Fanuc KAREL source: KT00935.KL

PROGRAM KT00935
%NOLOCKGROUP
VAR
  ENTRY: INTEGER
  PNAME: STRING[80]
  VNAME: STRING[80]
  STATUS: INTEGER
  VALUE: BOOLEAN
BEGIN
  ENTRY = 0
  PNAME = ''
  VNAME = 'VALUE'
  GET_VAR(ENTRY, PNAME, VNAME, VALUE, STATUS)
END KT00935
